(* CODESYS project Magazijn Overzetter Simulatie Structured Text 2V1.project
   Title: Simulatie Sorteer Station
   Author: Rene Potters/Gerard Harkema
   Version: 0.1.0
   Description: Simulatie voor opstelling Sorteer Station.
   Company: Avans

Project tree, tasks and I/O mapping:
  Device : EHV-CPU1025, Hitachi-IES, order no. EHV-CPU1025, version 3.5.4.11
      settings: IP Address = '192.168.1.31'
    application ApplicationSt
      libraries: Standard, * (System); Util, * (System); VisuDialogs, 3.5.16.40 (System)
      task MainTask (cyclic, interval t#20ms, priority 1) calls Main
      task Simulatie (cyclic, interval t#20ms, priority 1) calls MagazijnSim, OverzetterSim
    Basic : Basic, Hitachi-IES, version 3.4.4.0
      <Empty>
      <Empty>
      <Empty>
      <Empty>
      <Empty>
      <Empty>
      <Empty>
      <Empty>
      <Empty>
      <Empty>
      <Empty>
  Simulatie/
    program MagazijnSim [ST]
    global variables SIM
    program OverzetterSim [ST]
    data type OverzetterDUT
    data type MagazijnDUT
  text list GlobalTextList
  Programma Structured Text/
    function block OverzetterClass [ST]: initialize, cycle, isError, isKlaar, reset, start, noodstop
    function block StationClass [ST]: reset, isMagazijnLeeg, isError, isKlaar, start, cycle, initialize, noodstop
    function block MagazijnClass [ST]: initialize, cycle, start, isMagazijnLeeg, isError, reset, isKlaar, noodstop
    program Main [ST]
    TestProgramms/
      program MagazijnTest [ST]
      program OverzetterTest [ST]
    States/
      data type stationStates
      data type magazijnStates
      data type overzetterStates
    Structures/
      data type stationIO
      data type magazijnIO
      data type overzetterIO
      data type hmiIO
  global variables GVL
  Visualisaties/
    visualisation OverzetterHMI
    visualisation BekerMagazijnHMI
    visualisation StationHMI
*)

// Simulatie/OverzetterDUT
{attribute 'qualified_only'}
{attribute 'strict'}
TYPE OverzetterDUT :
(
	INHETMIDDEN, NAARRECHTS, ISRECHTS, NAARLINKS, ISLINKS, GEVALLEN
);
END_TYPE

// Programma Structured Text/Structures/stationIO
// Datum : 26 november 2026, Auteur: Gerard Harkema
TYPE stationIO :
STRUCT
	// IO van het magazijn
	magazijn		: magazijnIO;
	// IO van de overzetter
	overzetter		: overzetterIO;
END_STRUCT
END_TYPE

// Simulatie/MagazijnDUT
{attribute 'qualified_only'}
{attribute 'strict'}
TYPE MagazijnDUT :
(
	INGETROKKEN, INTREKKEN, UITGESTOTEN, UITSTOTEN, LEEG
);
END_TYPE

// Programma Structured Text/States/stationStates
// Datum : 26 november 2026, Auteur: Gerard Harkema
{attribute 'qualified_only'}
{attribute 'strict'}
TYPE stationStates :
(
	idle := 0,
	magazijn_uitstoten,
	wacht_magazijn_klaar,
	overzetten,
	wacht_overzetter_klaar,
	error
);
END_TYPE

// Programma Structured Text/States/magazijnStates
// Datum : 17 december 2020, Auteur: Gerard Harkema
{attribute 'qualified_only'}
{attribute 'strict'}
TYPE magazijnStates :
(
	idle := 0,
	in,
	travel_out,
	out,
	travel_in,
	error
);
END_TYPE

// Programma Structured Text/States/overzetterStates
// Datum : 17 december 2020, Auteur: Gerard Harkema
{attribute 'qualified_only'}
{attribute 'strict'}
TYPE overzetterStates :
(
	idle := 0,
	is_links,
	vaccuum_aanzetten,
	ga_naar_rechts,
	is_rechts,
	vaccuum_lossen,
	ga_naar_midden,
	is_midden,
	ga_naar_links,
	error
);
END_TYPE

// Programma Structured Text/Structures/magazijnIO
// Datum : 17 december 2020, Auteur: Gerard Harkema
TYPE magazijnIO :
STRUCT
	// Bekers magazijn zijn op
	Ix_MagazijnLeeg				: REFERENCE TO BOOL;
	// Beker is uit dekselmagazijn gestoten
	Ix_UitstoterBekerIn			: REFERENCE TO BOOL;
	// Uitstoter Beker haalt nieuwe beker op
	Ix_UitstoterBekerUit		: REFERENCE TO BOOL;
	// Beker uit magazijn stoten
	Qx_BekerUitstoten			: REFERENCE TO BOOL;

	//Perslucht is aanwezig
	Ix_PersluchtAanwezig 		: REFERENCE TO BOOL;

END_STRUCT
END_TYPE

// Programma Structured Text/Structures/overzetterIO
// Datum : 17 december 2020, Auteur: Gerard Harkema
TYPE overzetterIO :
STRUCT
	//Werkstuk door overzetter opgepakt
	Ix_VacuumAanwezig 		:REFERENCE TO BOOL;
	//Overzetter haalt beker op(linker pos.)
	Ix_OverzetterIsLinks 	:REFERENCE TO BOOL;
	//Overzetter plaatst beker op sorteerpositie
	Ix_OverzetterIsRechts 	:REFERENCE TO BOOL;
	//Beker aanwezig op detectiepositie
	
		//Beker oppakken
	Qx_VacuumAan 			:REFERENCE TO BOOL;
	//Beker loslaten
	Qx_BekerLossen 			:REFERENCE TO BOOL;
	//Overzetter naar bekermagazijn
	Qx_OverzetterLinks 		:REFERENCE TO BOOL;
	//Overzetter naar sorteerpositie
	Qx_OverzetterRechts 	:REFERENCE TO BOOL;

END_STRUCT
END_TYPE

// Programma Structured Text/Structures/hmiIO
// Datum : 17 december 2020, Auteur: Gerard Harkema
TYPE hmiIO :
STRUCT
	// Indrukken resetknop 
	Ix_Resetknop			: REFERENCE TO BOOL;
	// Keuzeknop staat op hand
	Ix_Hand					: REFERENCE TO BOOL;
	// Keuzeknop staat op auto
	Ix_Auto					: REFERENCE TO BOOL;
	// Indrukken noodstop
	Ix_Noodstop				: REFERENCE TO BOOL;
	// Bekers magazijn zijn op

	// Indrukken startknop
	Ix_Stopknop				: REFERENCE TO BOOL;
	// Indrukken stopknop
	Ix_Startknop			: REFERENCE TO BOOL;	
	//Perslucht is aanwezig

	// Visualisatie invisible Gele vlak
	Qx_GeleLamp				: REFERENCE TO BOOL;
	// Visualisatie invisible groene vlak
	Qx_GroeneLamp			: REFERENCE TO BOOL;
	// Visualisatie invisible rode vlak
	Qx_RodeLamp				: REFERENCE TO BOOL;

END_STRUCT
END_TYPE

// Simulatie/SIM
{attribute 'qualified_only'}
VAR_GLOBAL
	// Rotatie van de overzetter
	Vx_OvzRotate: INT := 0;
	// Visualisatie invisible blok
	Vx_OvzBlokLinks: BOOL := FALSE;
	// Visualisatie invisible blok
	Vx_OvzBlokOverzetter: BOOL := FALSE;
	// Visualisatie invisible blok
	Vx_OvzBlokRechts: BOOL := FALSE;
	// Visualisatie invisible blok
	Vx_OvzBlokGevallen: BOOL := FALSE;	
	// Magazijn opnieuw vullen (simulatie)
	Ix_MagazijnVullen 	: BOOL;
	// Simulatie visualisatie 
	Vw_Rotate45: INT := 45;
	// Visualisatie X positie van de uitstoter
	Vw_MagUitstoterBekerX: INT := 30;
	// Visualisatie invisible blok uitgestoten
	Vx_MagBlokUit: BOOL := TRUE;
	// Visualisatie invisible blok 1
	Vx_MagBlok1: BOOL := TRUE;
	// Visualisatie invisible blok 2
	Vx_MagBlok2: BOOL := TRUE;
	// Visualisatie invisible blok 3
	Vx_MagBlok3: BOOL := TRUE;
	// Visualisatie invisible blok 4
	Vx_MagBlok4: BOOL := TRUE;
	// Visualisatie invisible blokken
	Vx_MagBlok: ARRAY[1..8] OF BOOL;
	// Aantal blokken in het magazijn
	Vw_MagBlokAantal: INT := 4;
	// Simulatie onthoudt dat een blok maar 1x wordt uitgestoten
	Vw_MagBlok1X: INT := 0;
	// Simulatie error. Inverse logica.
	Vx_MagLuchtDrukError: BOOL := TRUE;
	// Simulatie error. Inverse logica.
	Vx_MagIsInError: BOOL := TRUE;
	// Simulatie error. Inverse logica.
	Vx_MagIsUitError: BOOL := TRUE;
	// Simulatie error. Inverse logica.
	Vx_OvzLuchtDrukError: BOOL := TRUE;
	// Simulatie error. Inverse logica.
	Vx_OvzIsLinksError: BOOL := TRUE;
	// Simulatie error. Inverse logica.
	Vx_OvzIsRechtsError: BOOL := TRUE;
	// Simulatie error. Inverse logica.
	Vx_OvzVacuumError: BOOL := TRUE;
	// Kleur van de blokken in het magazijn (lege plek = grijs)
	Vw_MagKleur: ARRAY[1..8] OF DWORD;
	// Kleur van het uitgestoten blok
	Vw_MagKleurUit: DWORD;
	// Kleur van het blok op de overzetter
	Vw_OvzKleur: DWORD := 16#FFC0C0C0;
	// Kleur van het blok dat klaarligt bij de uitgang van het magazijn
	Vw_MagKleurAfgifte: DWORD := 16#FFC0C0C0;
	// Er ligt een uitgestoten beker klaar bij de uitgang van het magazijn (voor de overzetter)
	Vx_MagBlokKlaar: BOOL := FALSE;
	// Afgifteplaats: kleur van de laatst afgegeven beker
	Vw_AfgifteKleur: DWORD := 16#FFA9A9A9;
	// Afgifteplaats: visualisatie invisible beker (inverse logica)
	Vx_AfgifteBeker: BOOL := TRUE;
	// Afgifteplaats: aantal afgegeven bekers
	Vi_AfgifteTeller: INT := 0;
	// Afgifteplaats leegmaken en teller op 0 (simulatie)
	Ix_AfgifteLegen: BOOL;
END_VAR

// GVL
VAR_GLOBAL
	// Indrukken resetknop 
	Ix_Resetknop: BOOL;
	// Keuzeknop staat op hand
	Ix_Hand: BOOL;
	// Keuzeknop staat op auto
	Ix_Auto: BOOL;
	// Indrukken noodstop
	Ix_Noodstop: BOOL;
	// Bekers magazijn zijn op
	Ix_MagazijnLeeg: BOOL;
	// Beker is uit dekselmagazijn gestoten
	Ix_UitstoterBekerIn: BOOL;
	// Uitstoter Beker haalt nieuwe beker op
	Ix_UitstoterBekerUit: BOOL;
	// Indrukken startknop
	Ix_Stopknop: BOOL := TRUE;
	// Indrukken stopknop
	Ix_Startknop: BOOL;	
	//Perslucht is aanwezig
	Ix_PersluchtAanwezig :BOOL;
	//Werkstuk door overzetter opgepakt
	Ix_VacuumAanwezig :BOOL;
	//Overzetter haalt beker op(linker pos.)
	Ix_OverzetterIsLinks :BOOL;
	//Overzetter plaatst beker op afgifteplaats
	Ix_OverzetterIsRechts :BOOL;
	// Beker uit magazijn stoten
	Qx_BekerUitstoten: BOOL;	
	//Beker oppakken
	Qx_VacuumAan :BOOL;
	//Beker loslaten
	Qx_BekerLossen :BOOL;
	//Overzetter naar bekermagazijn
	Qx_OverzetterLinks :BOOL;
	//Overzetter naar afgifteplaats
	Qx_OverzetterRechts :BOOL;
	// Visualisatie invisible Gele vlak
	Qx_GeleLamp: BOOL;
	// Visualisatie invisible groene vlak
	Qx_GroeneLamp: BOOL;
	// Visualisatie invisible rode vlak
	Qx_RodeLamp: BOOL;
	
END_VAR

// Programma Structured Text/Main
// Datum : 26 november 2026, Auteur: Gerard Harkema
// Main is het station: een magazijn en een overzetter, gecoordineerd door StationClass.
// Testen van een los object: vervang in de taakconfiguratie (MainTask) de aanroep van Main
// door MagazijnTest of OverzetterTest (map TestProgramms). De taak Simulatie blijft
// MagazijnSim en OverzetterSim aanroepen.
PROGRAM Main
VAR
	stationIO		: stationIO;
	station			: StationClass;
	initialized		: BOOL := FALSE;
END_VAR

IF NOT initialized THEN
	// Forceer perslucht aanwezig
	gvl.Ix_PersluchtAanwezig						:= TRUE;

	// ******** Magazijn ********/
	stationIO.magazijn.Ix_PersluchtAanwezig		REF= gvl.Ix_PersluchtAanwezig;
	stationIO.magazijn.Ix_MagazijnLeeg			REF= gvl.Ix_MagazijnLeeg;
	stationIO.magazijn.Ix_UitstoterBekerIn		REF= gvl.Ix_UitstoterBekerIn;
	stationIO.magazijn.Ix_UitstoterBekerUit		REF= gvl.Ix_UitstoterBekerUit;
	stationIO.magazijn.Qx_BekerUitstoten		REF= gvl.Qx_BekerUitstoten;

	// ******** Overzetter ********/
	//Werkstuk door overzetter opgepakt
	stationIO.overzetter.Ix_VacuumAanwezig		REF= gvl.Ix_VacuumAanwezig;
	//Overzetter haalt beker op (linker pos.)
	stationIO.overzetter.Ix_OverzetterIsLinks	REF= gvl.Ix_OverzetterIsLinks;
	//Overzetter plaatst beker op afgifteplaats (rechter pos.)
	stationIO.overzetter.Ix_OverzetterIsRechts	REF= gvl.Ix_OverzetterIsRechts;
	//Beker oppakken
	stationIO.overzetter.Qx_VacuumAan			REF= gvl.Qx_VacuumAan;
	//Beker loslaten
	stationIO.overzetter.Qx_BekerLossen			REF= gvl.Qx_BekerLossen;
	//Overzetter naar magazijn
	stationIO.overzetter.Qx_OverzetterLinks		REF= gvl.Qx_OverzetterLinks;
	//Overzetter naar afgifteplaats
	stationIO.overzetter.Qx_OverzetterRechts	REF= gvl.Qx_OverzetterRechts;

	station.initialize(stationIO);

	initialized := TRUE;
END_IF

// ******** Bediening ********/
IF gvl.Ix_Startknop THEN
	station.start();
	gvl.Ix_Startknop := FALSE;
END_IF

IF gvl.Ix_Noodstop THEN
	station.noodstop();
END_IF

IF gvl.Ix_Resetknop THEN
	station.reset();
END_IF

// ******** Signalering ********/
gvl.Qx_GroeneLamp	:= station.isKlaar();
gvl.Qx_RodeLamp		:= station.isError();
gvl.Qx_GeleLamp		:= station.isMagazijnLeeg();

station.cycle();

END_PROGRAM

// Programma Structured Text/StationClass
// Datum : 26 november 2026, Auteur: Gerard Harkema
// Station: coordineert een magazijn en een overzetter (compositie).
// De objecten praten alleen via methodes: start(), isKlaar(), isError().
FUNCTION_BLOCK StationClass
VAR
	IO				: REFERENCE TO stationIO;

	// ******** Magazijn ********/
	magazijn		: MagazijnClass;

	// ******** Overzetter ********/
	overzetter		: OverzetterClass;

	eState			: stationStates := stationStates.idle;
END_VAR

// Datum : 26 november 2026, Auteur: Gerard Harkema
METHOD reset
VAR_INPUT
END_VAR
// Reset geeft het station door aan beide objecten; die gaan eerst naar hun veilige stand
magazijn.reset();
overzetter.reset();
eState := stationStates.idle;
END_METHOD

// Datum : 26 november 2026, Auteur: Gerard Harkema
METHOD isMagazijnLeeg : BOOL
VAR_INPUT
END_VAR
isMagazijnLeeg := magazijn.isMagazijnLeeg();
END_METHOD

// Datum : 26 november 2026, Auteur: Gerard Harkema
METHOD isError : BOOL
VAR_INPUT
END_VAR
isError := (eState = stationStates.error);
END_METHOD

// Datum : 26 november 2026, Auteur: Gerard Harkema
METHOD isKlaar : BOOL
VAR_INPUT
END_VAR
isKlaar := (eState = stationStates.idle)
		AND magazijn.isKlaar()
		AND overzetter.isKlaar();
END_METHOD

// Datum : 26 november 2026, Auteur: Gerard Harkema
METHOD start : BOOL
VAR_INPUT
END_VAR
// Start een cyclus: een beker uit het magazijn naar de afgifteplaats.
// Kan alleen vanuit idle en als beide objecten in hun ruststand staan.
IF NOT isKlaar() THEN
	start := TRUE; // Failed (station blijft gewoon doorgaan met wat het deed)
	RETURN;
END_IF

eState := stationStates.magazijn_uitstoten;
start := FALSE; // oké
END_METHOD

// Datum : 26 november 2026, Auteur: Gerard Harkema
METHOD cycle
VAR
END_VAR
// Eerst de objecten
magazijn.cycle();
overzetter.cycle();

// Dan de fouten: een fout in een object zet het hele station in error
IF magazijn.isError() OR overzetter.isError() THEN
	eState := stationStates.error;
END_IF

// Dan de coordinatie, volgens het statediagram van StationClass
CASE eState OF
	stationStates.idle:
		; // wacht op start()

	stationStates.magazijn_uitstoten:
		IF magazijn.start() THEN		// TRUE = mislukt
			eState := stationStates.error;
		ELSE
			eState := stationStates.wacht_magazijn_klaar;
		END_IF

	stationStates.wacht_magazijn_klaar:
		IF magazijn.isKlaar() THEN
			eState := stationStates.overzetten;
		END_IF

	stationStates.overzetten:
		IF overzetter.start() THEN		// TRUE = mislukt
			eState := stationStates.error;
		ELSE
			eState := stationStates.wacht_overzetter_klaar;
		END_IF

	stationStates.wacht_overzetter_klaar:
		IF overzetter.isKlaar() THEN
			eState := stationStates.idle;
		END_IF

	stationStates.error:
		; // wacht op reset()
END_CASE
END_METHOD

// Datum : 26 november 2026, Auteur: Gerard Harkema
METHOD initialize
VAR_INPUT
	IORef			: REFERENCE TO stationIO;
END_VAR
IO REF= IORef;

// Elk object krijgt zijn eigen IO-structuur
magazijn.initialize(IO.magazijn);
overzetter.initialize(IO.overzetter);

eState := stationStates.idle;
END_METHOD

// Datum : 26 november 2026, Auteur: Gerard Harkema
METHOD noodstop
VAR_INPUT
END_VAR
// Noodstop geeft het station door aan beide objecten
magazijn.noodstop();
overzetter.noodstop();
eState := stationStates.error;
END_METHOD

END_FUNCTION_BLOCK

// Programma Structured Text/MagazijnClass
// Datum : 17 december 2020, Auteur: Gerard Harkema
FUNCTION_BLOCK MagazijnClass
VAR
	IO							: REFERENCE TO magazijnIO;

	xKlaar						: BOOL := FALSE;
	eState 						: magazijnStates := magazijnStates.idle;
END_VAR

// Datum : 17 december 2020, Auteur: Gerard Harkema
METHOD initialize
VAR_INPUT

	IORef		: REFERENCE TO magazijnIO;

END_VAR
IO 			REF= IORef;

eState 		:= magazijnStates.travel_in;
END_METHOD

// Datum : 17 december 2020, Auteur: Gerard Harkema
METHOD cycle
VAR_INPUT
END_VAR
CASE eState OF
	//magazijnStates.idle:
	//magazijnStates.in:
	magazijnStates.travel_out:
		IF IO.Ix_UitstoterBekerUit THEN
			eState 			:= magazijnStates.out;	
			IO.Qx_BekerUitstoten 	:= FALSE;
		END_IF
	magazijnStates.out:
		eState 				:= magazijnStates.travel_in;	
	magazijnStates.travel_in:
		IF IO.Ix_UitstoterBekerIn THEN
			eState 			:= magazijnStates.in;
			xKlaar			:= True;	
		END_IF
	
	//magazijnStates.error:
END_CASE
END_METHOD

// Datum : 17 december 2020, Auteur: Gerard Harkema
METHOD start : BOOL
VAR_INPUT
END_VAR
IF isMagazijnLeeg() THEN
	eState 				:= magazijnStates.error;
	IO.Qx_BekerUitstoten 	:= FALSE;
	start 		:= TRUE; // Failed
	RETURN;
END_IF

IF NOT IO.Ix_PersluchtAanwezig THEN
	eState 				:= magazijnStates.error;
	IO.Qx_BekerUitstoten 	:= FALSE;
	start 		:= TRUE; // Failed
	RETURN;
END_IF

IF NOT (eState = magazijnStates.in) THEN
	eState 				:= magazijnStates.error;
	IO.Qx_BekerUitstoten 	:= FALSE;
	start 		:= TRUE; // Failed
	RETURN;	
END_IF

xKlaar 					:= FALSE;
IO.Qx_BekerUitstoten 		:= TRUE;
eState 					:= magazijnStates.travel_out;

start 			:= FALSE; // oké
END_METHOD

// Datum : 17 december 2020, Auteur: Gerard Harkema
METHOD isMagazijnLeeg : BOOL
VAR_INPUT
END_VAR
isMagazijnLeeg := IO.Ix_MagazijnLeeg;
END_METHOD

// Datum : 17 december 2020, Auteur: Gerard Harkema
METHOD isError : BOOL
VAR_INPUT
END_VAR
isError := (eState = magazijnStates.error);
END_METHOD

// Datum : 17 december 2020, Auteur: Gerard Harkema
METHOD reset : BOOL
VAR_INPUT
END_VAR
eState 		:= magazijnStates.travel_in;
// Pas weer klaar als de ruststand bereikt is
xKlaar						:= FALSE;
END_METHOD

// Datum : 17 december 2020, Auteur: Gerard Harkema
METHOD isKlaar : BOOL
VAR_INPUT
END_VAR
isKlaar := xKlaar;
END_METHOD

// Datum : 17 december 2020, Auteur: Gerard Harkema
METHOD noodstop
VAR_INPUT
END_VAR
eState 				:= magazijnStates.error;
IO.Qx_BekerUitstoten 	:= FALSE;
END_METHOD

END_FUNCTION_BLOCK

// Programma Structured Text/OverzetterClass
// Datum : 17 december 2020, Auteur: Gerard Harkema
FUNCTION_BLOCK OverzetterClass
VAR
	IO							: reference to overzetterIO;

	xKlaar						: BOOL := FALSE;
	eState 						: overzetterStates := overzetterStates.idle;
	
	timer						: ton;
END_VAR

// Datum : 17 december 2020, Auteur: Gerard Harkema
METHOD initialize
VAR_INPUT
	IORef		: REFERENCE TO overzetterIO;
END_VAR
IO							REF= IORef;

IO.Qx_BekerLossen			:= FALSE;
IO.Qx_VacuumAan				:= FALSE;
IO.Qx_OverzetterLinks		:= FALSE;
IO.Qx_OverzetterRechts		:= TRUE;
eState 						:= overzetterStates.ga_naar_rechts;
END_METHOD

// Datum : 17 december 2020, Auteur: Gerard Harkema
METHOD cycle
VAR
END_VAR
CASE eState OF

//	overzetterStates.idle :
	overzetterStates.ga_naar_links:
		IF IO.Ix_OverzetterIsLinks THEN
			IO.Qx_OverzetterLinks 		:= FALSE;
			IO.Qx_VacuumAan 			:= TRUE;
			eState 					:= overzetterStates.is_links;
		END_IF;
	overzetterStates.is_links:
		IF IO.Ix_VacuumAanwezig THEN
			IO.Qx_OverzetterRechts 	:= TRUE;
			eState					:= overzetterStates.ga_naar_rechts;
	END_IF
//	overzetterStates.vaccuum_aanzetten:
	overzetterStates.ga_naar_rechts:
		IF IO.Ix_OverzetterIsRechts THEN
			IO.Qx_OverzetterRechts := FALSE;
			IO.Qx_VacuumAan 		:= FALSE;
			IO.Qx_BekerLossen 		:= TRUE;
			eState := overzetterStates.is_rechts;
		END_IF
	overzetterStates.is_rechts:
		IF NOT IO.Ix_VacuumAanwezig THEN
			IO.Qx_BekerLossen 		:= FALSE;
			IO.Qx_OverzetterLinks 	:= TRUE;
			eState 				:= overzetterStates.ga_naar_midden;
		END_IF
//	overzetterStates.vaccuum_lossen:
	overzetterStates.ga_naar_midden:
		IF timer.Q THEN
			IO.Qx_OverzetterLinks	:= FALSE;
			eState 				:= overzetterStates.is_midden;
			xKlaar 					:= TRUE;
		END_IF
		
	//overzetterStates.is_midden:
//	overzetterStates.error:
END_CASE

timer(IN:=(estate =overzetterStates.ga_naar_midden), PT:=T#2S);
END_METHOD

// Datum : 17 december 2020, Auteur: Gerard Harkema
METHOD isError : BOOL
VAR_INPUT
END_VAR
isError := (eState = overzetterStates.error);
END_METHOD

// Datum : 17 december 2020, Auteur: Gerard Harkema
METHOD isKlaar : BOOL
VAR_INPUT
END_VAR
isKlaar := xKlaar;
END_METHOD

// Datum : 17 december 2020, Auteur: Gerard Harkema
METHOD reset
VAR_INPUT
END_VAR
IO.Qx_BekerLossen			:= FALSE;
IO.Qx_VacuumAan				:= FALSE;
IO.Qx_OverzetterLinks		:= FALSE;
IO.Qx_OverzetterRechts		:= TRUE;
eState 						:= overzetterStates.ga_naar_rechts;
// Pas weer klaar als de ruststand bereikt is
xKlaar						:= FALSE;
END_METHOD

// Datum : 17 december 2020, Auteur: Gerard Harkema
METHOD start : BOOL
VAR_INPUT
END_VAR
IF NOT (eState = overzetterStates.is_midden) THEN
	eState 				:= overzetterStates.error;
//	IO.Qx_BekerUitstoten 	:= FALSE;
	start 	:= TRUE; // Failed
	RETURN;	
END_IF

xKlaar 					:= FALSE;
IO.Qx_OverzetterLinks 		:= TRUE;
eState 					:= overzetterStates.ga_naar_links;

start			:= FALSE; // oké
END_METHOD

// Datum : 17 december 2020, Auteur: Gerard Harkema
METHOD noodstop
VAR_INPUT
END_VAR
//Beker oppakken
IO.Qx_VacuumAan 			:=FALSE;
//Beker loslaten
IO.Qx_BekerLossen 			:=FALSE;
//Overzetter naar bekermagazijn
IO.Qx_OverzetterLinks 		:=FALSE;
//Overzetter naar sorteerpositie
IO.Qx_OverzetterRechts 	:=FALSE;

eState 				:= overzetterStates.error;
END_METHOD

END_FUNCTION_BLOCK

// Programma Structured Text/TestProgramms/MagazijnTest
// Datum : 17 december 2020, Auteur: Gerard Harkema
PROGRAM MagazijnTest
VAR
	xInitialaized				: BOOL := FALSE;
	
	magazijnIO					: magazijnIO;
	
	// Bekers magazijn zijn op
	Ix_MagazijnLeegRef			: REFERENCE TO BOOL;
	// Beker is uit dekselmagazijn gestoten
	Ix_UitstoterBekerInRef		: REFERENCE TO BOOL;
	// Uitstoter Beker haalt nieuwe beker op
	Ix_UitstoterBekerUitRef		: REFERENCE TO BOOL;
	// Beker uit magazijn stoten
	Qx_BekerUitstotenRef		: REFERENCE TO BOOL;
	
	magazijn: MagazijnClass;
	
END_VAR

IF NOT xInitialaized THEN

	// Forse Persluct aanwezig
	gvl.Ix_PersluchtAanwezig := TRUE;
	magazijnIO.Ix_PersluchtAanwezig		REF= gvl.Ix_PersluchtAanwezig;
	magazijnIO.Ix_MagazijnLeeg			REF= gvl.Ix_MagazijnLeeg;
	magazijnIO.Ix_UitstoterBekerIn 		REF= gvl.Ix_UitstoterBekerIn;
	magazijnIO.Ix_UitstoterBekerUit 	REF= gvl.Ix_UitstoterBekerUit;
	magazijnIO.Qx_BekerUitstoten 		REF= gvl.Qx_BekerUitstoten;

	magazijn.initialize(magazijnIO);

	xInitialaized	:= TRUE;
END_IF

IF Ix_Startknop THEN
	magazijn.start();
	Ix_Startknop := FALSE;
END_IF

IF Ix_Resetknop THEN
	magazijn.reset();
END_IF

IF Ix_Noodstop THEN
	magazijn.noodstop();
END_IF

Qx_GroeneLamp := magazijn.isKlaar();
Qx_RodeLamp := magazijn.isError();
Qx_GeleLamp := magazijn.isMagazijnLeeg();
 
magazijn.cycle();

END_PROGRAM

// Programma Structured Text/TestProgramms/OverzetterTest
// Datum : 17 december 2020, Auteur: Gerard Harkema
PROGRAM OverzetterTest
VAR
	xInitialaized				: BOOL := FALSE;

	overzetterIO				: overzetterIO;

	overzetter: OverzetterClass;
	
END_VAR

IF NOT xInitialaized THEN

	// Forse Persluct aanwezig
	gvl.Ix_PersluchtAanwezig := TRUE;
	
	//Werkstuk door overzetter opgepakt
	overzetterIO.Ix_VacuumAanwezig 		REF= gvl.Ix_VacuumAanwezig;
	//Overzetter haalt beker op(linker pos.)
	overzetterIO.Ix_OverzetterIsLinks 	REF= gvl.Ix_OverzetterIsLinks;
	//Overzetter plaatst beker op sorteerpositie
	overzetterIO.Ix_OverzetterIsRechts 	REF= gvl.Ix_OverzetterIsRechts;
	//Beker aanwezig op detectiepositie
	
		//Beker oppakken
	overzetterIO.Qx_VacuumAan 			REF= gvl.Qx_VacuumAan;
	//Beker loslaten
	overzetterIO.Qx_BekerLossen 			REF= gvl.Qx_BekerLossen;
	//Overzetter naar bekermagazijn
	overzetterIO.Qx_OverzetterLinks		REF= gvl.Qx_OverzetterLinks;
	//Overzetter naar sorteerpositie
	overzetterIO.Qx_OverzetterRechts 	REF= gvl.Qx_OverzetterRechts;

	overzetter.initialize(overzetterIO);

	xInitialaized	:= TRUE;
END_IF

IF Ix_Startknop THEN
	overzetter.start();
	Ix_Startknop := FALSE;
END_IF

IF Ix_Noodstop THEN
	overzetter.noodstop();
END_IF

IF Ix_Resetknop THEN
	overzetter.reset();
END_IF

Qx_GroeneLamp := overzetter.isKlaar();
Qx_RodeLamp := overzetter.isError();
 
overzetter.cycle();

END_PROGRAM

// Simulatie/MagazijnSim
PROGRAM MagazijnSim
VAR
	// Timer om uitstoten en intrekken te vertragen
	Fb_Pulse: BLINK;
	// Timer om intrekken te vertragen
	Fb_Trigger: F_TRIG;
	// Eerste keer om visualisatie te updaten
	Mx_FirstTime: BOOL := TRUE;
	// Afhandeling van het magazijn
	Me_MagState: MAGAZIJNDUT := MAGAZIJNDUT.INGETROKKEN;
	// Kleuren van de blokken in het magazijn, [1] = onderste (wordt als eerste uitgestoten)
	Mw_KleurRij: ARRAY[1..8] OF DWORD;
	// Hulpvariabelen voor het kiezen van een willekeurige kleur
	Mi_Indx: INT;
	Mu_Seed: UDINT := 1;
END_VAR
VAR CONSTANT
	// Metaal blank (zilver): metaal en reflecterend
	METAAL_BLANK: DWORD := 16#FFC0C0C0;
	// Metaal zwart (antraciet): metaal, niet reflecterend
	METAAL_ZWART: DWORD := 16#FF505050;
	// Kunststof rood: geen metaal, wel reflecterend
	KUNSTOF_ROOD: DWORD := 16#FFFF0000;
	// Kunststof zwart: geen metaal, niet reflecterend
	KUNSTOF_ZWART: DWORD := 16#FF000000;
	// Lege plek in het magazijn
	LEEG: DWORD := 16#FFA9A9A9;
END_VAR

//
// Common stuff.
//

IF (Mx_FirstTime) THEN
	SIM.Vw_MagBlokAantal := 8;
	SIM.Vx_MagBlokUit:= FALSE;
	
	// Vul het magazijn met blokken in willekeurige kleuren (materiaal + kleur).
	Mu_Seed := DINT_TO_UDINT(TIME_TO_DINT(TIME())) + Mu_Seed;
	FOR Mi_Indx := 1 TO 8 DO
		Mu_Seed := Mu_Seed * 1103515245 + 12345;
		CASE UDINT_TO_INT(SHR(Mu_Seed, 16) AND 3) OF
			0: Mw_KleurRij[Mi_Indx] := METAAL_BLANK;
			1: Mw_KleurRij[Mi_Indx] := METAAL_ZWART;
			2: Mw_KleurRij[Mi_Indx] := KUNSTOF_ROOD;
		ELSE
			Mw_KleurRij[Mi_Indx] := KUNSTOF_ZWART;
		END_CASE
	END_FOR
	Mx_FirstTime := FALSE;
END_IF

					
//
// Handle all pulse and trigger events.
//
Fb_Pulse(ENABLE:=TRUE,TIMELOW:=T#200MS, TIMEHIGH:=T#200MS);
Fb_Trigger(CLK:=Fb_Pulse.OUT);


//
// Only if no emergency active, start handling the simulation.
//
IF (SIM.Ix_MagazijnVullen) THEN
	Mx_FirstTime := TRUE;
	SIM.Ix_MagazijnVullen := FALSE;
	RETURN;
END_IF
	
//
// The pulse determines the speed of the cilinder to move in
// ore move out. The cilinder is only moved if the airpressure 
// is available.
//
IF (Fb_Trigger.Q AND SIM.Vx_MagLuchtDrukError) THEN
		
			
	CASE Me_MagState OF
		MAGAZIJNDUT.INGETROKKEN:
			IF (SIM.Vx_MagBlokUit) THEN
				SIM.Vw_MagBlokAantal := SIM.Vw_MagBlokAantal - 1;
				// Het onderste blok ligt nu klaar voor de overzetter; de rest zakt een plek.
				SIM.Vw_MagKleurAfgifte := Mw_KleurRij[1];
				SIM.Vx_MagBlokKlaar := TRUE;
				FOR Mi_Indx := 1 TO 7 DO
					Mw_KleurRij[Mi_Indx] := Mw_KleurRij[Mi_Indx + 1];
				END_FOR
				Mw_KleurRij[8] := LEEG;
			END_IF
		
			SIM.Vw_MagUitstoterBekerX := 1;
			SIM.Vw_MagBlok1X    	  := SIM.Vw_MagUitstoterBekerX;
			SIM.Vx_MagBlokUit         := FALSE;
	
			IF (Qx_BekerUitstoten) THEN
				Me_MagState := MAGAZIJNDUT.UITSTOTEN;
			END_IF

		MAGAZIJNDUT.INTREKKEN:
			SIM.Vw_MagUitstoterBekerX := SIM.Vw_MagUitstoterBekerX - 30;
			
			IF (SIM.Vw_MagUitstoterBekerX < 0) THEN 
				SIM.Vw_MagUitstoterBekerX := 0; 
			END_IF		
			
			IF (SIM.Vw_MagUitstoterBekerX = 0) THEN
				Me_MagState := MAGAZIJNDUT.INGETROKKEN;				
			END_IF		

			IF (Qx_BekerUitstoten) THEN
				Me_MagState := MAGAZIJNDUT.UITSTOTEN;
			END_IF	
	
		MAGAZIJNDUT.UITGESTOTEN:
			SIM.Vx_MagBlokUit         := SIM.Vx_MagBlok1;
						
			IF (NOT Qx_BekerUitstoten) THEN
				Me_MagState := MAGAZIJNDUT.INTREKKEN;
			END_IF	
		
		MAGAZIJNDUT.UITSTOTEN:
			SIM.Vw_MagUitstoterBekerX := SIM.Vw_MagUitstoterBekerX + 30;
			SIM.Vw_MagBlok1X    	  := SIM.Vw_MagUitstoterBekerX;			
		
			IF (SIM.Vw_MagUitstoterBekerX > 70) THEN
				Me_MagState := MAGAZIJNDUT.UITGESTOTEN;				
			END_IF		

			IF (NOT Qx_BekerUitstoten) THEN
				Me_MagState := MAGAZIJNDUT.INTREKKEN;
			END_IF	
		
	END_CASE

	GVL.Ix_UitstoterBekerIn  := (Me_MagState = MAGAZIJNDUT.INGETROKKEN) AND SIM.Vx_MagIsInError;
	GVL.Ix_UitstoterBekerUit := (Me_MagState = MAGAZIJNDUT.UITGESTOTEN) AND SIM.Vx_MagIsUitError;	
	GVL.Ix_MagazijnLeeg 	 := (SIM.Vw_MagBlokAantal <= 0) AND (Ix_UitstoterBekerIn);	
	
	SIM.Vx_MagBlok[8] := (SIM.Vw_MagBlokAantal >= 8);
	SIM.Vx_MagBlok[7] := (SIM.Vw_MagBlokAantal >= 7);
	SIM.Vx_MagBlok[6] := (SIM.Vw_MagBlokAantal >= 6);
	SIM.Vx_MagBlok[5] := (SIM.Vw_MagBlokAantal >= 5);		
	SIM.Vx_MagBlok[4] := (SIM.Vw_MagBlokAantal >= 4);
	SIM.Vx_MagBlok[3] := (SIM.Vw_MagBlokAantal >= 3);
	SIM.Vx_MagBlok[2] := (SIM.Vw_MagBlokAantal >= 2);
	SIM.Vx_MagBlok[1] := (SIM.Vw_MagBlokAantal >= 1);	

	// Kleur per plek voor de visualisatie
	FOR Mi_Indx := 1 TO 8 DO
		IF SIM.Vx_MagBlok[Mi_Indx] THEN
			SIM.Vw_MagKleur[Mi_Indx] := Mw_KleurRij[Mi_Indx];
		ELSE
			SIM.Vw_MagKleur[Mi_Indx] := LEEG;
		END_IF
	END_FOR
	IF SIM.Vx_MagBlokUit THEN
		SIM.Vw_MagKleurUit := Mw_KleurRij[1];
	ELSE
		SIM.Vw_MagKleurUit := LEEG;
	END_IF
	
END_IF

END_PROGRAM

// Simulatie/OverzetterSim
PROGRAM OverzetterSim
VAR
	// Timer om overzetten te vertragen
	Fb_Pulse: BLINK;
	// Timer om overzetten te vertragen
	Fb_Trigger: F_TRIG;
	// Eerste keer om visualisatie te updaten
	Mx_FirstTime: BOOL := TRUE;
	// Afhandeling van de overzetter
	Me_OvzState: OverzetterDUT := OVERZETTERDUT.INHETMIDDEN;	
	// Afhandeling van het blokje
	Me_BlokState: OverzetterDUT := OVERZETTERDUT.INHETMIDDEN;	
	// Duurt even voor het vacuum aanwezig is
	Mi_VacuumCntr: INT := 0;	
	// De overzetter heeft echt een beker vast (FALSE = leeg opgepakt, er lag niets klaar)
	Mx_MetBeker: BOOL := FALSE;
END_VAR
VAR CONSTANT


	// Inverse logica
	INVISABLE: BOOL := TRUE;
	// Inverse logica
	VISABLE: BOOL := FALSE;

END_VAR

// Initialisatie.

//
// Afgifteplaats leegmaken (knop in de visualisatie).
//
IF (SIM.Ix_AfgifteLegen) THEN
	SIM.Vi_AfgifteTeller := 0;
	SIM.Vx_AfgifteBeker  := INVISABLE;
	SIM.Vw_AfgifteKleur  := 16#FFA9A9A9;
	SIM.Ix_AfgifteLegen  := FALSE;
END_IF

IF (Mx_FirstTime) THEN
	Me_OvzState := OVERZETTERDUT.INHETMIDDEN;
	Me_BlokState := OVERZETTERDUT.ISLINKS;
	
	Mi_VacuumCntr := 0;
	Mx_MetBeker := FALSE;
	SIM.Vx_OvzRotate := 0;
	Mx_FirstTime := FALSE;
END_IF

//
// Afhandelen van de pulse events. Hierdoor loopt de simulatie los van de 
// TASK tijd.
//
Fb_Pulse(ENABLE:=TRUE,TIMELOW:=T#100MS, TIMEHIGH:=T#100MS);
Fb_Trigger(CLK:=Fb_Pulse.OUT);


//
// Only if no emergency active, start handling the simulation.
//
IF (GVL.Ix_Noodstop) THEN
	Mx_FirstTime := TRUE;	
	RETURN;
END_IF
	
//
// The pulse determines the speed of the cilinder to move in
// ore move out. The cilinder is only moved if the airpressure 
// is available.
//
IF (Fb_Trigger.Q AND SIM.Vx_OvzLuchtDrukError) THEN
	
	//
	// De status van de arm wordt los afgehandeld van het blokje. De beweging
	// van de arm staat hier namelijk helemaal los van.
	//
	
	CASE Me_OvzState OF
		
		OVERZETTERDUT.INHETMIDDEN:
			// 
			// De arm is in beweging naar links of naar rechts.
			// Indien de arm in de uiterste positie is wordt er van 
			// state gewisseld. Aangezien de arm in beweging is staan
			// de eindschakelaars uit.
			//
			
			IF (GVL.Qx_OverzetterLinks) THEN
				IF (SIM.Vx_OvzRotate > -90) THEN
					GVL.Ix_OverzetterIsLinks := FALSE;	
					GVL.Ix_OverzetterIsRechts := FALSE;			
					SIM.Vx_OvzRotate := SIM.Vx_OvzRotate - 10;
				ELSE
					Me_OvzState := OVERZETTERDUT.ISLINKS;			
				END_IF	
				
			END_IF
				 
			IF (GVL.Qx_OverzetterRechts) THEN
				IF (SIM.Vx_OvzRotate < 90) THEN
					GVL.Ix_OverzetterIsLinks := FALSE;	
					GVL.Ix_OverzetterIsRechts := FALSE;				
					SIM.Vx_OvzRotate := SIM.Vx_OvzRotate + 10;
				ELSE
					Me_OvzState := OVERZETTERDUT.ISRECHTS;				
				END_IF			
			END_IF
				
		OVERZETTERDUT.ISLINKS:
		    //
			// Arm staat in een uiterste stand. Eindschakelaar is ingeschakeld.
			// Zodra de arm weer wordt bewogen verandert de state.
			//
			
			GVL.Ix_OverzetterIsLinks := TRUE AND SIM.Vx_OvzIsLinksError;	

			IF (GVL.Qx_OverzetterRechts AND NOT GVL.Qx_OverzetterLinks) THEN
				GVL.Ix_OverzetterIsLinks := FALSE;				
				Me_OvzState := OVERZETTERDUT.INHETMIDDEN;		
			END_IF
			
		OVERZETTERDUT.ISRECHTS:
		    //
			// Arm staat in een uiterste stand. Eindschakelaar is ingeschakeld.
			// Zodra de arm weer wordt bewogen verandert de state.
			//
		
			GVL.Ix_OverzetterIsRechts := TRUE AND SIM.Vx_OvzIsRechtsError;	

			IF (GVL.Qx_OverzetterLinks AND NOT GVL.Qx_OverzetterRechts) THEN
				GVL.Ix_OverzetterIsRechts := FALSE;				
				Me_OvzState := OVERZETTERDUT.INHETMIDDEN;		
			END_IF			
			
		END_CASE

	END_IF	

	//
	// De status van het blokje hangt af van een aantal stuursignalen zoals waar
	// de arm zich bevindt, of er vacuum is en of er een beker lossen wordt gegeven.
	//
	
	CASE Me_BlokState OF
		OVERZETTERDUT.ISLINKS:
			//
			// Als de arm links is moet er eerst een vacuum opgebouwd worden alvorens het blokje 
			// opgepakt kan worden. Daarna verandert de state. Er ligt alleen een blokje links
			// als het magazijn er een heeft uitgestoten (SIM.Vx_MagBlokKlaar).
			//
			
			SIM.Vx_OvzBlokGevallen 	 := INVISABLE;
			SIM.Vx_OvzBlokLinks 	 := NOT SIM.Vx_MagBlokKlaar;
			SIM.Vx_OvzBlokOverzetter := INVISABLE;
			SIM.Vx_OvzBlokRechts 	 := INVISABLE;
			
			IF (GVL.Qx_VacuumAan AND SIM.Vx_OvzVacuumError AND GVL.Ix_OverzetterIsLinks) AND (NOT GVL.Qx_BekerLossen) THEN
				Mi_VacuumCntr := Mi_VacuumCntr + 1;
			END_IF
			
			IF (NOT GVL.Qx_VacuumAan AND SIM.Vx_OvzVacuumError) THEN
				Mi_VacuumCntr := 0;
			END_IF

			GVL.Ix_VacuumAanwezig := (Mi_VacuumCntr > 50);
	
			IF  ( GVL.Ix_VacuumAanwezig AND (Me_OvzState = OVERZETTERDUT.INHETMIDDEN)) THEN
				// Het blok wordt opgepakt en krijgt de kleur van het blok uit het magazijn.
				// Lag er geen blok klaar, dan beweegt de arm leeg (en komt er niets op de afgifteplaats).
				Mx_MetBeker := SIM.Vx_MagBlokKlaar;
				SIM.Vx_MagBlokKlaar := FALSE;
				SIM.Vw_OvzKleur := SIM.Vw_MagKleurAfgifte;
				Me_BlokState := OVERZETTERDUT.INHETMIDDEN;
			END_IF
			
		OVERZETTERDUT.INHETMIDDEN:
			//
			// Het blokje is in beweging zolang er vacuum is. Als er geen vacuum meer is
			// valt het blokje... Indien de arm helemaal rechts is kan het blokje gelost 
			// worden op de afgifteplaats. Dit moet met een Bekerlossen ondanks het feit dat er
			// geen vacuum meer is....
			//
			
			SIM.Vx_OvzBlokGevallen 	 := INVISABLE;
			SIM.Vx_OvzBlokLinks 	 := NOT SIM.Vx_MagBlokKlaar;
			SIM.Vx_OvzBlokOverzetter := NOT Mx_MetBeker;
			SIM.Vx_OvzBlokRechts 	 := INVISABLE;

		 	IF (GVL.Ix_OverzetterIsRechts) AND (NOT GVL.Qx_VacuumAan) AND (GVL.Qx_BekerLossen) THEN
				GVL.Ix_VacuumAanwezig := FALSE;
				IF Mx_MetBeker THEN
					// Beker komt op de afgifteplaats: zelfde kleur, teller omhoog.
					SIM.Vw_AfgifteKleur  := SIM.Vw_OvzKleur;
					SIM.Vx_AfgifteBeker  := VISABLE;
					SIM.Vi_AfgifteTeller := SIM.Vi_AfgifteTeller + 1;
				END_IF
				Me_BlokState := OVERZETTERDUT.ISRECHTS;		
				RETURN;		
			END_IF
			
			IF (NOT GVL.Ix_OverzetterIsRechts) AND (NOT GVL.Ix_OverzetterIsLinks) AND(NOT GVL.Qx_VacuumAan) THEN
				GVL.Ix_VacuumAanwezig := FALSE;
				Me_BlokState := OVERZETTERDUT.GEVALLEN;				
			END_IF

		OVERZETTERDUT.ISRECHTS:	
		    // 
			// Blokje is gelost op de afgifteplaats. Nu is het wachten tot de overzetter terug naar links wordt gestuurd.
			//
			
			SIM.Vx_OvzBlokGevallen 	 := INVISABLE;
			SIM.Vx_OvzBlokLinks 	 := NOT SIM.Vx_MagBlokKlaar;
			SIM.Vx_OvzBlokOverzetter := INVISABLE;
			SIM.Vx_OvzBlokRechts 	 := INVISABLE;
			
			IF (NOT GVL.Ix_OverzetterIsRechts) THEN
				Mx_MetBeker := FALSE;
				Me_BlokState := OVERZETTERDUT.ISLINKS;					
			END_IF

		OVERZETTERDUT.GEVALLEN:
			//
			// Blokje is gevallen..... Situatie herstelt zich zodra de arm helemaal links staat.
			//
				
			SIM.Vx_OvzBlokGevallen 	 := NOT Mx_MetBeker;
			SIM.Vx_OvzBlokLinks 	 := NOT SIM.Vx_MagBlokKlaar;
			SIM.Vx_OvzBlokOverzetter := INVISABLE;
			SIM.Vx_OvzBlokRechts 	 := INVISABLE;
			
			IF (GVL.Ix_OverzetterIsLinks) THEN
				Mx_MetBeker := FALSE;
				Me_BlokState := OVERZETTERDUT.ISLINKS;					
			END_IF				
	END_CASE

END_PROGRAM

// Visualisaties/OverzetterHMI
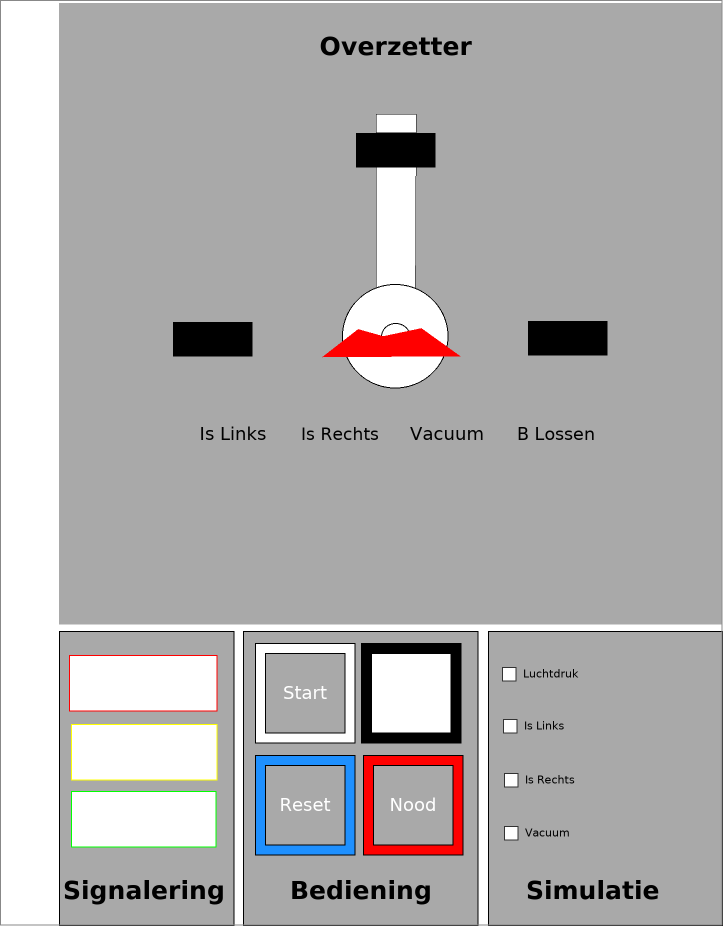
VISUALIZATION OverzetterHMI  // 723x926
    Rectangle (58,2 664x623)
    Polygon (233,394) (233,394) (273,434) (233,474) (193,434), "Is Links", colour toggle: Ix_OverzetterisLinks
    Polygon (340,394) (340,394) (380,434) (340,474) (300,434), "Is Rechts", colour toggle: Ix_OverzetterIsRechts
    Polygon (447,394) (447,394) (487,434) (447,474) (407,434), "Vacuum", colour toggle: Ix_VacuumAanwezig
    Polygon (376,131) (391,131) (416,131) (415,310) (376,310)
        p2858320360: SIM.Vx_OvzRotate
    Polygon (556,394) (556,394) (596,434) (556,474) (516,434), "B Lossen", colour toggle: Qx_BekerLossen
    Polygon (376,114) (391,114) (416,114) (416,132) (376,132), colour toggle: Qx_VacuumAan
        p2858320360: SIM.Vx_OvzRotate
    Polygon (356,133) (371,133) (435,133) (435,167) (356,167), invisible if: SIM.Vx_OvzBlokOverzetter, colour variable: SIM.Vw_OvzKleur
        p2277200375: SIM.Vx_OvzRotate
    Polygon (173,322) (188,322) (252,322) (252,356) (173,356), invisible if: SIM.Vx_OvzBlokLinks, colour variable: SIM.Vw_MagKleurAfgifte
    Polygon (528,321) (543,321) (607,321) (607,355) (528,355), invisible if: SIM.Vx_AfgifteBeker, colour variable: SIM.Vw_AfgifteKleur
    Ellipse (342,284 106x104)
    Ellipse (381,323 29x27)
    Polygon (358,329) (383,336) (421,328) (460,356) (322,357), invisible if: SIM.Vx_OvzBlokGevallen, colour variable: SIM.Vw_OvzKleur
        p2277200375: SIM.Vx_OvzRotate
    Label (294,31 204x30), "Overzetter"
    Group (59,631 175x295)
        Rectangle (0,0 175x295)
        Rectangle (10,24 148x56), colour toggle: Qx_RodeLamp
        Rectangle (12,93 146x56), colour toggle: Qx_GeleLamp
        Rectangle (12,160 145x56), colour toggle: Qx_GroeneLamp
        Label (10,236 150x46), "Signalering"
    Group (243,631 235x295)
        Rectangle (0,0 235x295)
        Group (12,12 100x100)
            RoundedRectangle (0,0 100x100)
            RoundedRectangle (10,10 80x80), "Start", tooltip "Start knop", colour toggle: Ix_Startknop
                OnMouseDown: execute { Ix_Startknop := TRUE; }
                OnMouseUp: execute { Ix_Startknop := FALSE; }
        Group (118,12 100x100)
            RoundedRectangle (0,0 100x100)
            RoundedRectangle (10,10 80x80), "Stop", tooltip "Stop knop", colour toggle: Ix_Stopknop
                OnMouseDown: execute { Ix_Stopknop := FALSE; }
                OnMouseUp: execute { Ix_Stopknop := TRUE; }
        Group (12,124 100x100)
            RoundedRectangle (0,0 100x100)
            RoundedRectangle (10,10 80x80), "Reset", tooltip "Reset knop", colour toggle: Ix_Resetknop
                OnMouseDown: execute { Ix_Resetknop := TRUE; }
                OnMouseUp: execute { Ix_Resetknop := FALSE; }
        Group (120,124 100x100)
            RoundedRectangle (0,0 100x100), "Nood"
            RoundedRectangle (10,10 80x80), "Nood", tooltip "Noodstop", colour toggle: Ix_Noodstop
                OnMouseDown: execute { Ix_Noodstop := NOT Ix_Noodstop; }
        Label (43,236 150x46), "Bediening"
    Group (488,631 235x295)
        Group (0,0 235x295)
            Rectangle (0,0 235x295)
            Label (30,236 150x46), "Simulatie"
        Checkbox (12,17 196x52), "Luchtdruk", variable: SIM.Vx_OvzLuchtDrukError
        Checkbox (13,69 196x52), "Is Links", variable: SIM.Vx_OvzIsLinksError
        Checkbox (14,123 196x52), "Is Rechts", variable: SIM.Vx_OvzIsRechtsError
        Checkbox (14,176 196x52), "Vacuum", variable: SIM.Vx_OvzVacuumError
END_VISUALIZATION

// Visualisaties/BekerMagazijnHMI
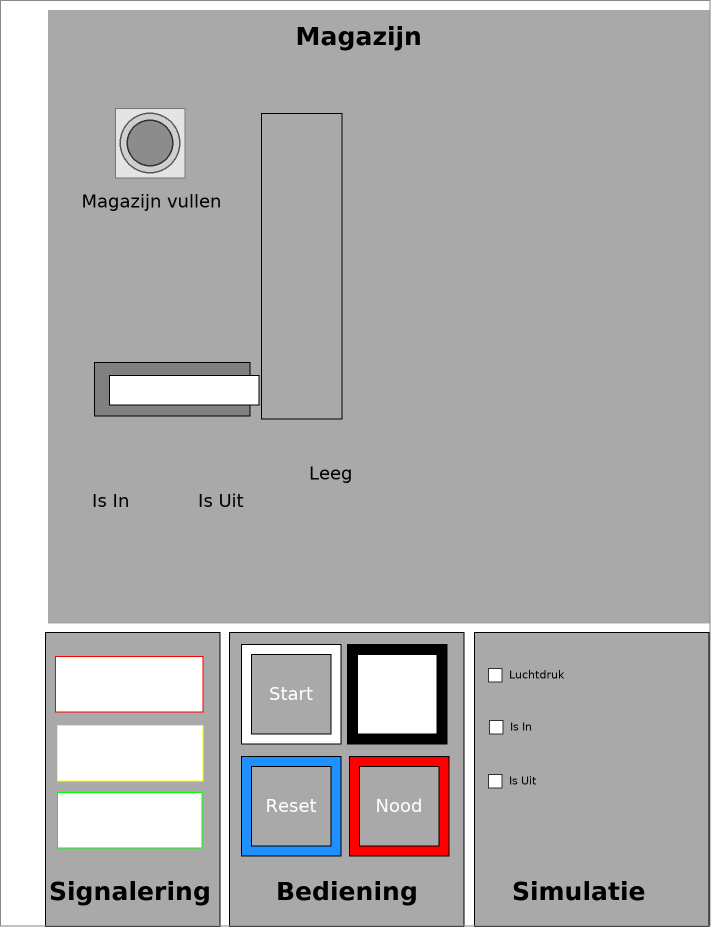
VISUALIZATION BekerMagazijnHMI  // 711x927
    Rectangle (47,9 664x615)
    Polygon (286,461) (316,461) (346,461) (376,461) (331,541), "Leeg", colour toggle: Ix_MagazijnLeeg
    Polygon (111,461) (111,461) (151,501) (111,541) (71,501), "Is In", colour toggle: Ix_UitstoterBekerIn
    Polygon (221,461) (221,461) (261,501) (221,541) (181,501), "Is Uit", colour toggle: Ix_UitstoterBekerUit
    Rectangle (94,362 156x54)
    Rectangle (261,113 81x306)
    Rectangle (353,376 61x29), colour variable: SIM.Vw_MagKleurUit
    Rectangle (266,341 61x29), colour variable: SIM.Vw_MagKleur[2]
    Rectangle (266,305 61x29), colour variable: SIM.Vw_MagKleur[3]
    Rectangle (266,269 61x29), colour variable: SIM.Vw_MagKleur[4]
    Rectangle (266,376 61x29), colour variable: SIM.Vw_MagKleur[1]
        p3560616238: SIM.Vw_MagBlok1X
    Rectangle (109,375 150x30)
        p3560616238: SIM.Vw_MagUitstoterBekerX
    Label (284,21 150x30), "Magazijn"
    Group (45,632 664x295)
        Group (0,0 664x295)
            Group (429,0 235x295)
                Rectangle (0,0 235x295)
                Label (30,236 150x46), "Simulatie"
            Group (0,0 175x295)
                Rectangle (0,0 175x295)
                Rectangle (10,24 148x56), colour toggle: Qx_RodeLamp
                Rectangle (12,93 146x56), colour toggle: Qx_GeleLamp
                Rectangle (12,160 145x56), colour toggle: Qx_GroeneLamp
                Label (10,236 150x46), "Signalering"
            Group (184,0 235x295)
                Rectangle (0,0 235x295)
                Group (12,12 100x100)
                    RoundedRectangle (0,0 100x100)
                    RoundedRectangle (10,10 80x80), "Start", tooltip "Start knop", colour toggle: Ix_Startknop
                        OnMouseDown: execute { Ix_Startknop := TRUE; }
                        OnMouseUp: execute { Ix_Startknop := FALSE; }
                Group (118,12 100x100)
                    RoundedRectangle (0,0 100x100)
                    RoundedRectangle (10,10 80x80), "Stop", tooltip "Stop knop", colour toggle: Ix_Stopknop
                        OnMouseDown: execute { Ix_Stopknop := FALSE; }
                        OnMouseUp: execute { Ix_Stopknop := TRUE; }
                Group (12,124 100x100)
                    RoundedRectangle (0,0 100x100)
                    RoundedRectangle (10,10 80x80), "Reset", tooltip "Reset knop", colour toggle: Ix_Resetknop
                        OnMouseDown: execute { Ix_Resetknop := TRUE; }
                        OnMouseUp: execute { Ix_Resetknop := FALSE; }
                Group (120,124 100x100)
                    RoundedRectangle (0,0 100x100), "Nood"
                    RoundedRectangle (10,10 80x80), "Nood", tooltip "Noodstop", colour toggle: Ix_Noodstop
                        OnMouseDown: execute { Ix_Noodstop := NOT Ix_Noodstop; }
                Label (43,236 150x46), "Bediening"
        Checkbox (441,17 196x52), "Luchtdruk", variable: SIM.Vx_MagLuchtDrukError
        Checkbox (442,69 196x52), "Is In", variable: SIM.Vx_MagIsInError
        Checkbox (441,123 196x52), "Is Uit", variable: SIM.Vx_MagIsUitError
    Rectangle (266,197 61x29), colour variable: SIM.Vw_MagKleur[6]
    Rectangle (266,161 61x29), colour variable: SIM.Vw_MagKleur[7]
    Rectangle (266,125 61x29), colour variable: SIM.Vw_MagKleur[8]
    Rectangle (266,232 61x29), colour variable: SIM.Vw_MagKleur[5]
    Polygon (74,189) (104,189) (134,189) (229,203) (129,217), "Magazijn vullen", colour toggle: Ix_MagazijnLeeg
    PushSwitch (115,108 70x70), tooltip "Magazijn vullen", variable: SIM.Ix_MagazijnVullen, behaviour: TOGGLE, style: Switch-PushSwitch-Gray
END_VISUALIZATION

// Visualisaties/StationHMI
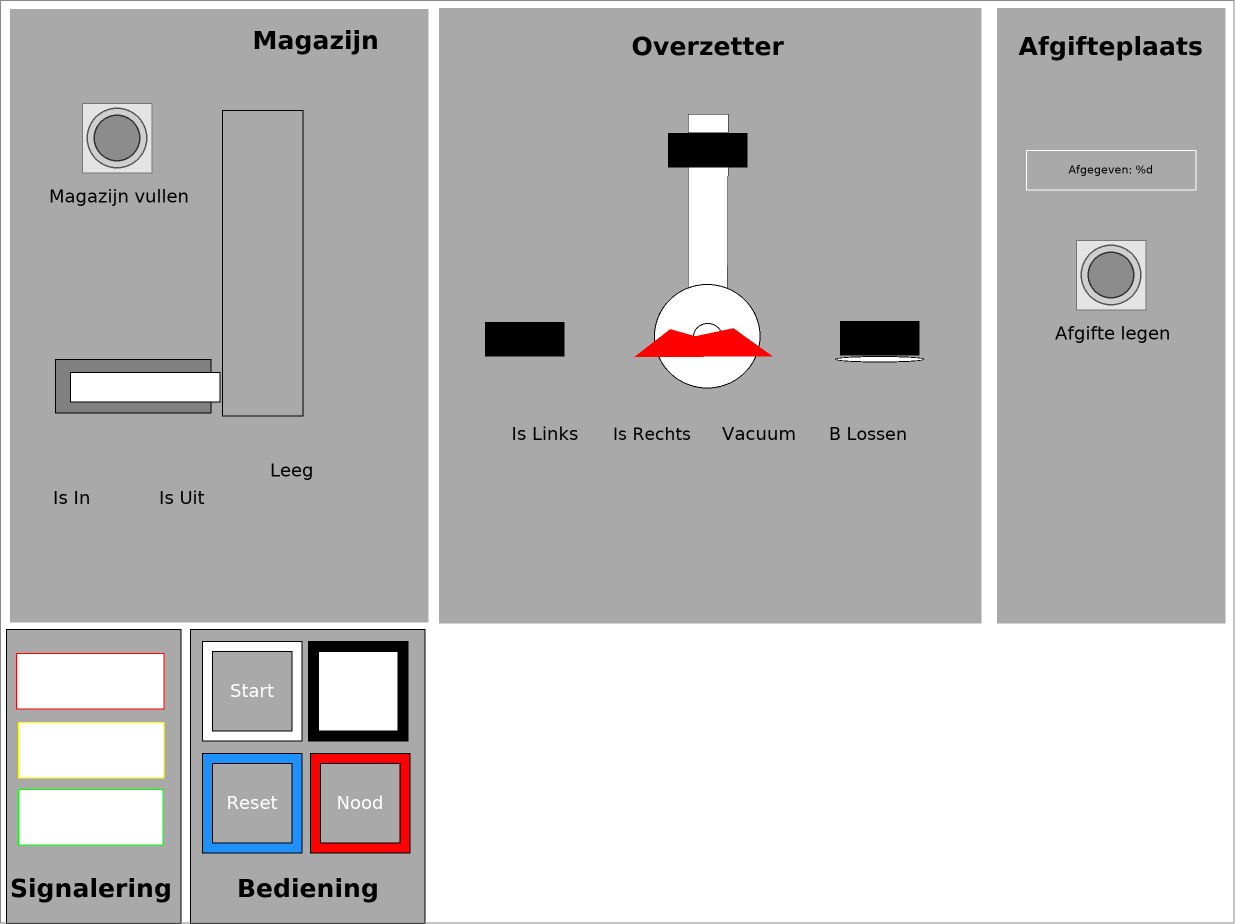
VISUALIZATION StationHMI  // 1235x924
    Rectangle (9,8 420x615)
    Polygon (247,458) (277,458) (307,458) (337,458) (292,538), "Leeg", colour toggle: Ix_MagazijnLeeg
    Polygon (72,458) (72,458) (112,498) (72,538) (32,498), "Is In", colour toggle: Ix_UitstoterBekerIn
    Polygon (182,458) (182,458) (222,498) (182,538) (142,498), "Is Uit", colour toggle: Ix_UitstoterBekerUit
    Rectangle (55,359 156x54)
    Rectangle (222,110 81x306)
    Rectangle (314,373 61x29), colour variable: SIM.Vw_MagKleurUit
    Rectangle (227,338 61x29), colour variable: SIM.Vw_MagKleur[2]
    Rectangle (227,302 61x29), colour variable: SIM.Vw_MagKleur[3]
    Rectangle (227,266 61x29), colour variable: SIM.Vw_MagKleur[4]
    Rectangle (227,373 61x29), colour variable: SIM.Vw_MagKleur[1]
        p3560616238: SIM.Vw_MagBlok1X
    Rectangle (70,372 150x30)
        p3560616238: SIM.Vw_MagUitstoterBekerX
    Label (241,25 150x30), "Magazijn"
    Group (6,629 175x295)
        Rectangle (0,0 175x295)
        Rectangle (10,24 148x56), colour toggle: Qx_RodeLamp
        Rectangle (12,93 146x56), colour toggle: Qx_GeleLamp
        Rectangle (12,160 145x56), colour toggle: Qx_GroeneLamp
        Label (10,236 150x46), "Signalering"
    Group (190,629 235x295)
        Rectangle (0,0 235x295)
        Group (12,12 100x100)
            RoundedRectangle (0,0 100x100)
            RoundedRectangle (10,10 80x80), "Start", tooltip "Start knop", colour toggle: Ix_Startknop
                OnMouseDown: execute { Ix_Startknop := TRUE; }
                OnMouseUp: execute { Ix_Startknop := FALSE; }
        Group (118,12 100x100)
            RoundedRectangle (0,0 100x100)
            RoundedRectangle (10,10 80x80), "Stop", tooltip "Stop knop", colour toggle: Ix_Stopknop
                OnMouseDown: execute { Ix_Stopknop := FALSE; }
                OnMouseUp: execute { Ix_Stopknop := TRUE; }
        Group (12,124 100x100)
            RoundedRectangle (0,0 100x100)
            RoundedRectangle (10,10 80x80), "Reset", tooltip "Reset knop", colour toggle: Ix_Resetknop
                OnMouseDown: execute { Ix_Resetknop := TRUE; }
                OnMouseUp: execute { Ix_Resetknop := FALSE; }
        Group (120,124 100x100)
            RoundedRectangle (0,0 100x100), "Nood"
            RoundedRectangle (10,10 80x80), "Nood", tooltip "Noodstop", colour toggle: Ix_Noodstop
                OnMouseDown: execute { Ix_Noodstop := NOT Ix_Noodstop; }
        Label (43,236 150x46), "Bediening"
    Rectangle (227,194 61x29), colour variable: SIM.Vw_MagKleur[6]
    Rectangle (227,158 61x29), colour variable: SIM.Vw_MagKleur[7]
    Rectangle (227,122 61x29), colour variable: SIM.Vw_MagKleur[8]
    Rectangle (227,229 61x29), colour variable: SIM.Vw_MagKleur[5]
    Rectangle (438,7 544x617)
    Polygon (545,394) (545,394) (585,434) (545,474) (505,434), "Is Links", colour toggle: Ix_OverzetterisLinks
    Polygon (652,394) (652,394) (692,434) (652,474) (612,434), "Is Rechts", colour toggle: Ix_OverzetterIsRechts
    Polygon (759,394) (759,394) (799,434) (759,474) (719,434), "Vacuum", colour toggle: Ix_VacuumAanwezig
    Polygon (688,131) (703,131) (728,131) (727,310) (688,310)
        p2858320360: SIM.Vx_OvzRotate
    Polygon (868,394) (868,394) (908,434) (868,474) (828,434), "B Lossen", colour toggle: Qx_BekerLossen
    Polygon (688,114) (703,114) (728,114) (728,132) (688,132), colour toggle: Qx_VacuumAan
        p2858320360: SIM.Vx_OvzRotate
    Polygon (668,133) (683,133) (747,133) (747,167) (668,167), invisible if: SIM.Vx_OvzBlokOverzetter, colour variable: SIM.Vw_OvzKleur
        p2277200375: SIM.Vx_OvzRotate
    Polygon (485,322) (500,322) (564,322) (564,356) (485,356), invisible if: SIM.Vx_OvzBlokLinks, colour variable: SIM.Vw_MagKleurAfgifte
    Polygon (840,321) (855,321) (919,321) (919,355) (840,355), invisible if: SIM.Vx_AfgifteBeker, colour variable: SIM.Vw_AfgifteKleur
    Ellipse (654,284 106x104)
    Ellipse (693,323 29x27)
    Polygon (670,329) (695,336) (733,328) (772,356) (634,357), invisible if: SIM.Vx_OvzBlokGevallen, colour variable: SIM.Vw_OvzKleur
        p2277200375: SIM.Vx_OvzRotate
    Label (606,31 204x30), "Overzetter"
    PushSwitch (82,103 70x70), tooltip "Magazijn vullen", variable: SIM.Ix_MagazijnVullen, behaviour: TOGGLE, style: Switch-PushSwitch-Gray
    Polygon (41,184) (71,184) (101,184) (197,196) (96,212), "Magazijn vullen"
    Rectangle (996,7 230x617)
    Label (1009,31 204x30), "Afgifteplaats"
    Rectangle (1026,150 170x40), "Afgegeven: %d", text variable: SIM.Vi_AfgifteTeller
    PushSwitch (1076,240 70x70), tooltip "Afgifte legen", variable: SIM.Ix_AfgifteLegen, behaviour: TOGGLE, style: Switch-PushSwitch-Gray
    Polygon (1035,321) (1065,321) (1095,321) (1191,333) (1090,349), "Afgifte legen"
    Ellipse (835,356 89x6)
END_VISUALIZATION
